(* IEC 61131-3 sources: Test-Git_ESME26/TestProgettoESME_26.fbsproj/AxisModule_Migration_Example.device.xml.v3^/Plc Logic.plclogic.xml.v3^/Application.application.xml.v3^/Sercos_AxisModule/WriteIDN, 1 file *)

(* ---- FC_SercosWriteIDN.fn.st ---- *)
FUNCTION FC_SercosWriteIDN : DINT
VAR_INPUT
	i_uiTopoAddr : UINT;
	i_etSercosParameterType : ET_SercosParameterType;
	i_uiIDN : UINT;
	i_etWriteIDNType : ET_SercosWriteIDNType;
	i_dwValue : DWORD;
END_VAR
VAR
	dwIDN : DWORD;
	dwValue : DWORD;
END_VAR

dwValue := i_dwValue;

IF i_etSercosParameterType = ET_SercosParameterType.S_Parameter THEN
	dwIDN := i_uiIDN;
ELSE
	dwIDN := 16#8000 + i_uiIDN;
END_IF

FC_SercosWriteIDN := SMM6xx.FC_SercosWriteServiceDataByTopAddr(
	i_wTopoAddr := i_uiTopoAddr,
	i_dwIDN := dwIDN,
	i_wType := TO_UINT(i_etWriteIDNType),
	i_lwPointerToData := TO_LWORD(ADR(dwValue)),
	i_wMaxDataLen := 2);
